PROGRAM MAIN
VAR
END_VAR

PRG_IO_In();
PRG_Seq();
PRG_IO_Out();

END_PROGRAM

(* stored: Version 1.1.0.1
   POU MAIN: Id {4c0e654f-7d72-4b04-b772-7a5f16f12ddb}, SpecialFunc None *)
